(* IEC 61131-3 sources: plcassist-cli/packages/volt-lsp-iec/test-corpus/lenze-mid/Device/Plc Logic/Application/Library Manager/L_DCO_DriveCommunication, 14 files *)

(* ---- GETBOOLEANPROPERTY.fun ---- *)
FUNCTION GETBOOLEANPROPERTY : BOOL
VAR_INPUT
	STKEY : WSTRING;
END_VAR
END_FUNCTION

(* ---- GETCOMPANY.fun ---- *)
FUNCTION GETCOMPANY : WSTRING
END_FUNCTION

(* ---- GETNUMBERPROPERTY.fun ---- *)
FUNCTION GETNUMBERPROPERTY : DINT
VAR_INPUT
	STKEY : WSTRING;
END_VAR
END_FUNCTION

(* ---- GETTEXTPROPERTY.fun ---- *)
FUNCTION GETTEXTPROPERTY : WSTRING
VAR_INPUT
	STKEY : WSTRING;
END_VAR
END_FUNCTION

(* ---- GETTEXTPROPERTY2.fun ---- *)
FUNCTION GETTEXTPROPERTY2 : POINTER TO WSTRING
VAR_INPUT
	STKEY : WSTRING;
END_VAR
END_FUNCTION

(* ---- GETTITLE.fun ---- *)
FUNCTION GETTITLE : WSTRING
END_FUNCTION

(* ---- GETVERSION.fun ---- *)
FUNCTION GETVERSION : VERSION
END_FUNCTION

(* ---- GETVERSIONPROPERTY.fun ---- *)
FUNCTION GETVERSIONPROPERTY : VERSION
VAR_INPUT
	STKEY : WSTRING;
END_VAR
END_FUNCTION

(* ---- GLOBALTEXTLIST.fb ---- *)
FUNCTION_BLOCK GLOBALTEXTLIST
VAR
	M_TEXTLISTFILE : STRING(255);
	_STNAMESPACE : STRING;
END_VAR
END_FUNCTION_BLOCK

(* ---- L_DCO_AXIS_REF_BASE.fb ---- *)
FUNCTION_BLOCK L_DCO_AXIS_REF_BASE EXTENDS IoDrvBase
VAR_INPUT
	UDITIMEOUT : UDINT := 10000;
	USICHANNEL : USINT := 1;
	ASDOREADDATA : ARRAY [1..c_wSdoMaxNumTotal] OF L_DCO_SdoData;
	ASDOWRITEDATA : ARRAY [1..c_wSdoMaxNumTotal] OF L_DCO_SdoData;
END_VAR
VAR_OUTPUT
	UIDEVICEID : UINT := 0;
	UINETID : UINT := 0;
	XCOMMUNICATIONOK : BOOL := FALSE;
	ECOMMUNICATIONSTATE : L_DCO_CommState := 0;
	AXISNAME : STRING := '';
END_VAR
VAR
	DWAXISID : DWORD;
	AXISINSTANCE : __XWORD;
	READIDX : DWORD := 1;
	WRITEIDX : DWORD := 1;
	M_PSLAVECONNECTOR : POINTER TO IoConfigConnector;
	M_PAXISCONNECTOR : POINTER TO IoConfigConnector;
	M_IIODRV : ICmpIoDrv;
	M_IIODRVPARAMETER : ICmpIoDrvParameter;
	XCOPYDATA : BOOL := TRUE;
	SINSTANCESTR : STRING;
	XPARACCESSBYSEMANOTSUPPORTED : BOOL := TRUE;
	DWSEMAPARREADACCESS : DWORD;
	DWSEMAPARWRITEACCESS : DWORD;
	C_WSDOMAXNUMTOTAL : WORD := 10;
	C_WSDOMAXNUM : WORD := 5;
	WMAXSDONUMBERREAD : WORD;
	WMAXSDONUMBERREADTOTAL : WORD;
	WMAXSDONUMBERWRITE : WORD;
	WMAXSDONUMBERWRITETOTAL : WORD;
END_VAR
END_FUNCTION_BLOCK

METHOD GETAXISSLOT : UINT
END_METHOD

METHOD GETREADPARAMETERCONTAINER : POINTER TO L_DCO_SDOData
END_METHOD

METHOD GETWRITEPARAMETERCONTAINER : POINTER TO L_DCO_SDOData
END_METHOD

METHOD INITIALIZE : UDINT
VAR_INPUT
	WMODULETYPE : UINT;
	DWINSTANCE : UDINT;
	PCONNECTOR : POINTER TO IoConfigConnector;
END_VAR
END_METHOD

METHOD IODRVREADPARAMETER : UDINT
VAR_INPUT
	PCONNECTOR : POINTER TO IoConfigConnector;
	PPARAMETER : POINTER TO IoConfigParameter;
	PDATA : POINTER TO BYTE;
	DWBITSIZE : DWORD;
	DWBITOFFSET : DWORD;
END_VAR
END_METHOD

METHOD IODRVWRITEPARAMETER : UDINT
VAR_INPUT
	PCONNECTOR : POINTER TO IoConfigConnector;
	PPARAMETER : POINTER TO IoConfigParameter;
	PDATA : POINTER TO BYTE;
	DWBITSIZE : DWORD;
	DWBITOFFSET : DWORD;
END_VAR
END_METHOD

METHOD QUERYINTERFACE : POINTER TO POINTER TO BYTE
VAR_INPUT
	IID : DWORD;
	PRESULT : POINTER TO UDINT;
END_VAR
END_METHOD

METHOD FB_INIT : BOOL
VAR_INPUT
	BINITRETAINS : BOOL;
	BINCOPYCODE : BOOL;
END_VAR
END_METHOD

(* ---- L_DCO_READDRIVEPARAMETER.fb ---- *)
FUNCTION_BLOCK L_DCO_READDRIVEPARAMETER
VAR_INPUT
	XEXECUTE : BOOL := FALSE;
	WINDEX : WORD := 0;
	BYSUBINDEX : BYTE := 0;
	XUSEINDEXASPARAM : BOOL := FALSE;
END_VAR
VAR_OUTPUT
	XDONE : BOOL := FALSE;
	XBUSY : BOOL := FALSE;
	XERROR : BOOL := FALSE;
	EERROR : L_DCO_Error := L_DCO_Error.L_DCO_No_Error;
	DWDATA : DWORD := 0;
	BYNROFBYTE : BYTE := 0;
END_VAR
VAR_IN_OUT
	AXIS : L_DCO_AXIS_REF_BASE;
END_VAR
VAR
	IDX : DWORD;
	XEXECUTEOLD : BOOL;
	SDOREAD : POINTER TO L_DCO_SdoData;
	SDOMAXREADNUM : WORD;
	SAXISNAME : STRING;
	SDOREADINTERNAL : BOOL := FALSE;
	SDONUMSTART : WORD;
	SDONUMEND : WORD;
	AXISINSTANCE : __XWORD := 0;
	XRESETOUTPUTS : BOOL;
	ABORT : BOOL;
	SDOACCESSAXISREF : BOOL;
END_VAR
END_FUNCTION_BLOCK

(* ---- L_DCO_READDRIVEPARAMETERSTRING.fb ---- *)
FUNCTION_BLOCK L_DCO_READDRIVEPARAMETERSTRING
VAR_INPUT
	XEXECUTE : BOOL := FALSE;
	WINDEX : WORD := 0;
	BYSUBINDEX : BYTE := 0;
	XUSEINDEXASPARAM : BOOL := FALSE;
END_VAR
VAR_OUTPUT
	XDONE : BOOL := FALSE;
	XBUSY : BOOL := FALSE;
	XERROR : BOOL := FALSE;
	EERROR : L_DCO_Error := L_DCO_Error.L_DCO_No_Error;
	SVALUE : STRING(255) := '';
	BYNROFBYTE : BYTE := 0;
END_VAR
VAR_IN_OUT
	AXIS : L_DCO_AXIS_REF_BASE;
END_VAR
VAR
	IDX : DWORD;
	XSEMASUPPORTEDBYAXIS : BOOL;
	XEXECUTEOLD : BOOL;
	XSEMASUPPORT : BOOL;
	SDOREAD : POINTER TO L_DCO_SdoData;
	SDONUMSTART : WORD;
	SDONUMEND : WORD;
	SDOREADINTERNAL : BOOL := FALSE;
	AXISINSTANCE : __XWORD := 0;
	SVALUEINT : STRING(255) := '';
	SAXISNAME : STRING;
	XRESETOUTPUTS : BOOL;
	ABORT : BOOL;
	SDOACCESSAXISREF : BOOL;
END_VAR
END_FUNCTION_BLOCK

(* ---- L_DCO_TRANSFERDRIVEPARAMETER.fb ---- *)
FUNCTION_BLOCK L_DCO_TRANSFERDRIVEPARAMETER
VAR_INPUT
	XEXECUTE : BOOL := FALSE;
	PSCPARAMETERDATA : POINTER TO L_DCO_TranferData;
	DWSIZEPARAMETERDATA : DWORD := 0;
	XUSEINDEXASPARAM : BOOL := FALSE;
END_VAR
VAR_OUTPUT
	XDONE : BOOL := FALSE;
	XBUSY : BOOL := FALSE;
	XERROR : BOOL := FALSE;
	EERROR : L_DCO_Error := L_DCO_Error.L_DCO_No_Error;
	WINDEXCOUNTER : WORD := 0;
END_VAR
VAR_IN_OUT
	AXIS : L_DCO_AXIS_REF_BASE;
END_VAR
VAR
	L_DCO_READDRIVEPARAMETER1 : L_DCO_ReadDriveParameter;
	L_DCO_WRITEDRIVEPARAMETER1 : L_DCO_WriteDriveParameter;
	IDX : DWORD;
	WSTEP : WORD;
	DWADRESSCOUNTER : DWORD;
	DWARRAYSIZE : DWORD;
	PSCPARAMETERDATAINTERN : POINTER TO L_DCO_TranferData;
	SCDUMMY : L_DCO_TranferData;
	DWSINGLESIZE : DWORD;
	AXISINSTANCE : __XWORD := 0;
	SAXISNAME : STRING;
END_VAR
END_FUNCTION_BLOCK

(* ---- L_DCO_WRITEDRIVEPARAMETER.fb ---- *)
FUNCTION_BLOCK L_DCO_WRITEDRIVEPARAMETER
VAR_INPUT
	XEXECUTE : BOOL := FALSE;
	WINDEX : WORD := 0;
	BYSUBINDEX : BYTE := 0;
	XUSEINDEXASPARAM : BOOL := FALSE;
	DWDATA : DWORD := 0;
	BYNROFBYTE : BYTE := 4;
END_VAR
VAR_OUTPUT
	XDONE : BOOL := FALSE;
	XBUSY : BOOL := FALSE;
	XERROR : BOOL := FALSE;
	EERROR : L_DCO_Error := L_DCO_Error.L_DCO_No_Error;
END_VAR
VAR_IN_OUT
	AXIS : L_DCO_AXIS_REF_BASE;
END_VAR
VAR
	IDX : DWORD;
	XEXECUTEOLD : BOOL;
	SDOWRITE : POINTER TO L_DCO_SdoData;
	SAXISNAME : STRING;
	SDOWRITEINTERNAL : BOOL := FALSE;
	SDONUMSTART : WORD;
	SDONUMEND : WORD;
	AXISINSTANCE : __XWORD := 0;
	XRESETOUTPUTS : BOOL;
	ABORT : BOOL;
	SDOACCESSAXISREF : BOOL;
END_VAR
END_FUNCTION_BLOCK
